Fanuc KAREL source: kb00094.KL

PROGRAM KB00094
%STACKSIZE=65535
%PRIORITY=65535
%NOLOCKGROUP
VAR
P1 : INTEGER
BEGIN
P1=1
GET_TIME(P1)
END KB00094
